(* IEC 61131-3 sources: kns-pump-station/src/POUs/Station/FB_Ats, 2 files *)

(* ---- FB_Ats.decl.st ---- *)
// Назначение: АВР насосов (04 §9): отказ насоса, у которого был запрос в прошлом цикле (Fault —
//             нет ОС пуска, авария ПЧ, пропадание ОС; или блокировка станции насоса axTrip —
//             недогрузка, перегрев), — насос снят АВР до возврата доступности (KNS1.ATS),
//             событие 101006 с номером насоса, получившего новый запрос в окне STN_ATS_WINDOW.
//             Смена режима оператором, пропадание напряжения и сухой ход станции — не АВР. Условия
//             «недостаточно насосов» (KNS1.LACK) и «нет резерва» (KNS1.NORES); их задержки — в Cfg
//             тревог, подавления — в ядре станции (FB_StationCore).
// Автор:      kr0nsch
// Версия:     0.1.0
// Документ:   docs/DESIGN.md, раздел 6.6; docs/04_algorithms.md, раздел 9
FUNCTION_BLOCK FB_Ats
VAR_INPUT
    xEnable     : BOOL;             // станция в «Автомате»
    aitfPump    : ARRAY[1..GVL_Const.STN_PUMP_COUNT] OF PL.I_MotorVfd;
    axRun       : ARRAY[1..GVL_Const.STN_PUMP_COUNT] OF BOOL;   // запросы этого цикла (FB_PumpRotation)
    axTrip      : ARRAY[1..GVL_Const.STN_PUMP_COUNT] OF BOOL;   // блокировка станции насоса: недогрузка, перегрев
    uiRequired  : UINT;
    uiAvailable : UINT;
    uiForeign   : UINT;
    itfTime     : PL.I_TimeSource;
    itfEvents   : I_StationEventSink;
END_VAR
VAR_IN_OUT CONSTANT
    stCfg : ST_StationCfg;          // uiDutyMax
END_VAR
VAR_OUTPUT
    xAtsActive  : BOOL;             // есть насос, снятый АВР и ещё недоступный (KNS1.ATS)
    axRemoved   : ARRAY[1..GVL_Const.STN_PUMP_COUNT] OF BOOL;
    xLack       : BOOL;             // uiRequired > uiAvailable + uiForeign (KNS1.LACK; задержка — в Cfg тревоги)
    xNoReserve  : BOOL;             // uiAvailable < MIN(uiDutyMax, STN_DUTY_MAX) + 1 (KNS1.NORES; подавления — в ядре)
    udiAtsCount : UDINT;            // АВР с запуска (HMI)
END_VAR
VAR
    axRunPrev  : ARRAY[1..GVL_Const.STN_PUMP_COUNT] OF BOOL;    // запросы прошлого цикла
    xWindow    : BOOL;              // идёт окно поиска замены (событие 101006)
    axReqAtAts : ARRAY[1..GVL_Const.STN_PUMP_COUNT] OF BOOL;    // запросы в момент АВР: замена — новый запрос
    fbWindow   : PL.FB_Delay;       // окно STN_ATS_WINDOW
END_VAR
VAR_TEMP
    uiPump    : UINT;               // номер насоса
    xFailed   : BOOL;               // насос с запросом отказал в этом цикле
    xAvail    : BOOL;               // насос доступен
    xFault    : BOOL;               // отказ насоса (Fault) или фиксация станции (axTrip)
    uiNewPump : UINT;               // насос, получивший новый запрос в окне
END_VAR

(* ---- FB_Ats.impl.st ---- *)
// 1. Отказ запрошенного насоса (запрос был в прошлом цикле): Fault или фиксация станции
xFailed := FALSE;
FOR uiPump := 1 TO GVL_Const.STN_PUMP_COUNT DO
    xAvail := FALSE;
    xFault := FALSE;
    IF aitfPump[uiPump] <> 0 THEN
        xAvail := aitfPump[uiPump].Available;
        xFault := aitfPump[uiPump].Fault;
    END_IF
    xFault := xFault OR axTrip[uiPump];
    IF xEnable AND axRunPrev[uiPump] AND NOT axRemoved[uiPump] AND xFault THEN
        axRemoved[uiPump] := TRUE;
        udiAtsCount := udiAtsCount + 1;
        xFailed := TRUE;
    END_IF
    // насос снят АВР, пока снова не станет доступен — сброшен и в Auto (04 §9.1). Фиксация станции
    // действует на устройство только с его вызова, поэтому без отказа и фиксации, а не только Available
    IF axRemoved[uiPump] AND xAvail AND NOT xFault THEN
        axRemoved[uiPump] := FALSE;
    END_IF
END_FOR

// 2. Окно поиска замены: новый запрос насоса, которого не было в момент отказа (FB_PumpRotation
//    назначает замену в том же цикле, если резерв готов). Снятый АВР насос заменой не бывает: при
//    блокировке станции (недогрузка, перегрев) он ещё доступен и запрошен в цикле отказа
IF xFailed THEN
    xWindow := TRUE;
    fbWindow.Preset(xValue := FALSE);
    FOR uiPump := 1 TO GVL_Const.STN_PUMP_COUNT DO
        axReqAtAts[uiPump] := axRunPrev[uiPump] AND NOT axRemoved[uiPump];
    END_FOR
END_IF
fbWindow(xIn := xWindow, tOnDelay := GVL_Const.STN_ATS_WINDOW, itfTime := itfTime);
IF xWindow THEN
    uiNewPump := 0;
    FOR uiPump := 1 TO GVL_Const.STN_PUMP_COUNT DO
        IF uiNewPump = 0 AND axRun[uiPump] AND NOT axReqAtAts[uiPump] AND NOT axRemoved[uiPump] THEN
            uiNewPump := uiPump;
        END_IF
    END_FOR
    IF uiNewPump <> 0 THEN
        xWindow := FALSE;
        IF itfEvents <> 0 THEN
            itfEvents.LogEvent(eEvent := E_StationEvent.AtsPumpIn, rValue := UINT_TO_REAL(uiNewPump));
        END_IF
    ELSIF fbWindow.xOut OR NOT xEnable THEN
        xWindow := FALSE;                               // заменить нечем: KNS1.LACK по своему условию
    END_IF
END_IF

// 3. Сводные условия
xAtsActive := FALSE;
FOR uiPump := 1 TO GVL_Const.STN_PUMP_COUNT DO
    xAtsActive := xAtsActive OR axRemoved[uiPump];
    axRunPrev[uiPump] := axRun[uiPump];
END_FOR
xLack := uiRequired > uiAvailable + uiForeign;
// резерв — сверх насосов обычного режима: ступенчатое и ПИД работают не больше чем MIN(uiDutyMax, STN_DUTY_MAX)
xNoReserve := uiAvailable < MIN(stCfg.uiDutyMax, GVL_Const.STN_DUTY_MAX) + 1;
